(* IEC 61131-3 sources: virtual-bottling-plant/plc/src/packml, 3 files *)

(* ---- PackMLHasStarted.st ---- *)
(* TRUE once a machine has left Idle on its way to production (running, waiting or held). *)
FUNCTION PackMLHasStarted : BOOL
  VAR_INPUT
    State : E_PackMLState;
  END_VAR
  PackMLHasStarted := State = PML_STARTING OR State = PML_EXECUTE OR State = PML_SUSPENDING
                      OR State = PML_SUSPENDED OR State = PML_UNSUSPENDING
                      OR State = PML_HOLDING OR State = PML_HELD OR State = PML_UNHOLDING;
END_FUNCTION

(* ---- FB_PackagingUnit.st ---- *)
(* What every packaging machine has in common: PackML, merged line/HMI commands, debounced
   blocked/starved, and Admin.StopReason (PLC-13). Machine FBs add their own causes and
   setpoints. *)
FUNCTION_BLOCK FB_PackagingUnit
  VAR_INPUT
    LineCmd : ST_MachineCmd;   (* from FB_LineSequencer *)
    OwnCmd : E_Command;        (* from the bridge, this machine only *)
    StopReasonCmd : INT;       (* operator reason code from the HMI, 0 = none *)
    HoldId : INT;              (* first active alarm of this machine, 0 = none *)
    LineHoldId : INT;          (* line alarm that holds every machine, 0 = none *)
    Blocked : BOOL;            (* raw: output conveyor full *)
    Starved : BOOL;            (* raw: no input and nothing coming (upstream not producing) *)
    StarvedDelayMs : UDINT;
    Running : BOOL;
    NowMs : UDINT;
  END_VAR
  VAR_OUTPUT
    Status : ST_PackagingStatus;
    RunOut : BOOL;
  END_VAR
  VAR
    PackML : FB_PackML;
    BlockedDelay : FB_SimTon;
    StarvedDelay : FB_SimTon;
    Cmd : ST_MachineCmd;
    LastState : E_PackMLState;
  END_VAR
  VAR CONSTANT
    BLOCKED_DELAY_MS : UDINT := 2000;
  END_VAR

  BlockedDelay(IN := Blocked, PT := BLOCKED_DELAY_MS, NowMs := NowMs);
  StarvedDelay(IN := Starved, PT := StarvedDelayMs, NowMs := NowMs);

  Cmd.Start := LineCmd.Start OR OwnCmd = CMD_START;
  Cmd.Stop := LineCmd.Stop OR OwnCmd = CMD_STOP;
  Cmd.Reset := LineCmd.Reset OR OwnCmd = CMD_RESET;
  Cmd.Abort := LineCmd.Abort OR OwnCmd = CMD_ABORT;
  Cmd.Clear := LineCmd.Clear OR OwnCmd = CMD_CLEAR;

  PackML(Cmd := Cmd, HoldCause := HoldId <> 0 OR LineHoldId <> 0,
         SuspendCause := BlockedDelay.Q OR StarvedDelay.Q, Running := Running, NowMs := NowMs);

  (* StopReason: cleared when production resumes, set automatically to the alarm id on a
     hold (1-99), overwritten by the operator's reason code from the HMI (>= 100). *)
  IF PackML.State = PML_EXECUTE AND LastState <> PML_EXECUTE THEN
    Status.StopReason := 0;
  END_IF;
  IF (PackML.State = PML_HOLDING OR PackML.State = PML_HELD) AND Status.StopReason = 0 THEN
    IF HoldId <> 0 THEN
      Status.StopReason := HoldId;
    ELSE
      Status.StopReason := LineHoldId;
    END_IF;
  END_IF;
  IF StopReasonCmd <> 0 THEN
    Status.StopReason := StopReasonCmd;
  END_IF;
  LastState := PackML.State;

  Status.State := PackML.State;
  Status.Mode := MODE_PRODUCTION;
  Status.Blocked := BlockedDelay.Q;
  Status.Starved := StarvedDelay.Q;
  RunOut := PackML.RunOut;
END_FUNCTION_BLOCK

(* ---- FB_PackML.st ---- *)
(* PackML state machine (PLC-01, ISA-TR88.00.02), shared by every packaging machine.
   Acting states (Starting, Holding, Stopping...) complete on the motor feedback, or after
   FEEDBACK_TIMEOUT_MS so a missing feedback can never lock the machine in a transition. *)
FUNCTION_BLOCK FB_PackML
  VAR_INPUT
    Cmd : ST_MachineCmd;     (* one-scan commands *)
    HoldCause : BOOL;        (* internal fault: jam, breakdown, material out, comms (PLC-10) *)
    SuspendCause : BOOL;     (* external: blocked or starved (PLC-10) *)
    Running : BOOL;          (* motor running feedback *)
    NowMs : UDINT;
  END_VAR
  VAR_OUTPUT
    State : E_PackMLState := PML_STOPPED;
    RunOut : BOOL;           (* motor run command *)
  END_VAR
  VAR
    InState : FB_SimTon;
    LastState : E_PackMLState := PML_STOPPED;
  END_VAR
  VAR CONSTANT
    FEEDBACK_TIMEOUT_MS : UDINT := 5000;
  END_VAR

  InState(IN := TRUE, PT := FEEDBACK_TIMEOUT_MS, NowMs := NowMs);

  IF Cmd.Abort AND State <> PML_ABORTING AND State <> PML_ABORTED THEN
    State := PML_ABORTING;
  END_IF;

  CASE State OF
    PML_ABORTING:
      IF NOT Running OR InState.Q THEN State := PML_ABORTED; END_IF;
    PML_ABORTED:
      IF Cmd.Clear THEN State := PML_CLEARING; END_IF;
    PML_CLEARING:
      State := PML_STOPPED;
    PML_STOPPED:
      IF Cmd.Reset THEN State := PML_RESETTING; END_IF;
    PML_RESETTING:
      State := PML_IDLE;
    PML_IDLE:
      IF Cmd.Stop THEN
        State := PML_STOPPING;
      ELSIF Cmd.Start AND NOT HoldCause THEN
        State := PML_STARTING;
      END_IF;
    PML_STARTING, PML_UNHOLDING:
      IF Cmd.Stop THEN
        State := PML_STOPPING;
      ELSIF HoldCause THEN
        State := PML_HOLDING;
      ELSIF Running OR InState.Q THEN
        State := PML_EXECUTE;
      END_IF;
    PML_EXECUTE:
      IF Cmd.Stop THEN
        State := PML_STOPPING;
      ELSIF HoldCause THEN
        State := PML_HOLDING;
      ELSIF SuspendCause THEN
        State := PML_SUSPENDING;
      END_IF;
    PML_SUSPENDING:
      State := PML_SUSPENDED;
    PML_SUSPENDED:
      IF Cmd.Stop THEN
        State := PML_STOPPING;
      ELSIF HoldCause THEN
        State := PML_HOLDING;
      ELSIF NOT SuspendCause THEN
        State := PML_UNSUSPENDING;
      END_IF;
    PML_UNSUSPENDING:
      State := PML_EXECUTE;
    PML_HOLDING:
      IF NOT Running OR InState.Q THEN State := PML_HELD; END_IF;
    PML_HELD:
      IF Cmd.Stop THEN
        State := PML_STOPPING;
      ELSIF Cmd.Reset AND NOT HoldCause THEN
        State := PML_UNHOLDING;
      END_IF;
    PML_STOPPING:
      IF NOT Running OR InState.Q THEN State := PML_STOPPED; END_IF;
    PML_COMPLETE:
      IF Cmd.Reset THEN State := PML_RESETTING; END_IF;
  ELSE
    State := PML_STOPPED;
  END_CASE;

  IF State <> LastState THEN
    LastState := State;
    InState(IN := FALSE, PT := FEEDBACK_TIMEOUT_MS, NowMs := NowMs);
  END_IF;

  (* Suspended keeps the motor on: the machine waits for bottles or room and resumes by itself *)
  RunOut := State = PML_STARTING OR State = PML_EXECUTE OR State = PML_SUSPENDING
            OR State = PML_SUSPENDED OR State = PML_UNSUSPENDING OR State = PML_UNHOLDING;
END_FUNCTION_BLOCK
